Staubli VAL3: click_refreshIOMsg.pgx

program click_refreshIOMsg()
begin
  nMsgType=3
  call initMsg()
  call rs:getLog(sRobotMsg,nMsgType)
  userPageSet("message","btnAllMsg","style.backgroundColor","#FFFFFF")
  userPageSet("message","btnRobotMsg","style.backgroundColor","#FFFFFF")
  userPageSet("message","btnTrajMsg","style.backgroundColor","#FFFFFF")
  userPageSet("message","btnIOMsg","style.backgroundColor","#33FF33")
end
